Fanuc KAREL source: KB00114.KL

PROGRAM KB00114
%NOLOCKGROUP
%ENVIRONMENT KCLOP
VAR
  P1: STRING[80]
  P2: INTEGER
BEGIN
  P1 = 'A'
  P2 = 1
  KCL_NO_WAIT(P1, P2)
END KB00114
